//============================================================
// 文件: PLC_Logic.scl
// 项目: PLC-Robot-Integration-Demo (PLC控制ABB机器人码垛)
// 平台: TIA Portal V16+ / S7-1214C DC/DC/DC
// 内容: 伺服控制FB / 主顺控FB / 故障处理FB / 急停处理
// 版本: V2.3  日期: 2026-09-02
// 变更: V1.0 基础正反转+限位保护
//       V2.0 增加完整顺控、故障码、急停安全处理
//       V2.1 超时改锁存+定时器卫生(修超时后无法复位/误超时)
//            故障灯无故障时强制熄灭; 启动命令改600ms脉冲式;
//            满垛输出qRobotReset(DI2)通知机器人清垛位计数
//       V2.2 定时器实例声明由IEC_TIMER改为TON多重实例(IEC_TIMER是
//            定时器背景SDT, 不能按FB方式直接调用, "从源生成块"编译报错);
//            故障复位不再清nParts——机器人侧nCount(PERS)仅在满垛DI2时
//            清零, 两侧计数必须同步保持, 否则中垛复位后垛位错位且
//            PLC等满垛/机器人等DI2互等死锁
//       V2.3 bHomeDone/nParts/nPallet移入VAR RETAIN: 掉电重启后PLC侧
//            计数不再清零, 与机器人nCount(PERS)断电保持对齐, 堵住
//            断电重启失步入口(VAR RETAIN为IEC 61131-3标准声明段)
//============================================================
//
// ----------------- I/O 交叉引用表(调试用) -----------------
// I0.0 启动SB1(常开)      I0.1 停止SB2(常闭)
// I0.2 复位SB3            I0.3 手动/自动旋钮(自动=1)
// I0.4 正限位SQ1          I0.5 反限位SQ2
// I0.6 机器人"允许抓取"DO1 I0.7 物料检测光电E3Z
// I1.0 急停回路反馈(常闭)  I1.1 安全门开关(常闭)
// I1.2 机器人"码垛完成"DO2 I1.3 机器人故障DO3
// I1.4 伺服报警ALM(断=报警) I1.5 伺服就绪RDY
// Q0.0 脉冲PUL+  Q0.4 方向DIR+  Q0.3 伺服使能KA1
// Q0.1 运行绿灯 Q0.2 报警红灯  Q0.5 蜂鸣器    Q0.6 待机黄灯
// Q0.7 机器人DI1启动  Q1.0 机器人DI2复位
// MW10 电流  MW12 电压  MW14 温度  MW16 计数  MW22 故障码
// ----------------------------------------------------------
//============================================================

//============================================================
// 块1: FB_ServoCtrl —— 伺服使能/点动/限位保护/报警锁存
//============================================================
FUNCTION_BLOCK "FB_ServoCtrl"
{ S7_Optimized_Access := 'TRUE' }
VERSION: 1.0

VAR_INPUT
    bPowerOn    : BOOL;    // 使能命令(来自顺控或手动)
    bReset      : BOOL;    // 报警复位
    bJogFwd     : BOOL;    // 手动点动正转
    bJogRev     : BOOL;    // 手动点动反转
    bFwdLimit   : BOOL;    // 正向限位SQ1(1=压合)
    bRevLimit   : BOOL;    // 反向限位SQ2(1=压合)
    bServoReady : BOOL;    // 驱动器RDY(1=就绪)
    bServoFault : BOOL;    // 驱动器ALM(1=报警, 现场常闭取反后送入)
    bEStopOK    : BOOL;    // 急停回路(1=正常)
END_VAR

VAR_OUTPUT
    qEnable     : BOOL;    // 伺服使能 -> KA1 -> CN1.DI1(SON)
    qFwdAllow   : BOOL;    // 允许正转(软件许可)
    qRevAllow   : BOOL;    // 允许反转(软件许可)
    qRun        : BOOL;    // 运行中标志
    qAlarm      : BOOL;    // 伺服报警锁存输出
END_VAR

VAR
    bFaultLock  : BOOL;    // 故障锁存位
    iDiag       : INT;     // 诊断码(供HMI显示)
END_VAR

BEGIN
    //---- 1) 故障锁存: 报警或急停立即置位 ----
    IF bServoFault OR NOT bEStopOK THEN
        bFaultLock := TRUE;
        iDiag := 16#0101;              // 伺服报警/急停类
    END_IF;

    //---- 2) 双限位同时压合 = 接线故障, 同样锁存 ----
    IF bFwdLimit AND bRevLimit THEN
        bFaultLock := TRUE;
        iDiag := 16#0102;
    END_IF;

    //---- 3) 复位: 故障源消失后按复位才解锁 ----
    IF bReset AND NOT bServoFault AND bEStopOK
       AND NOT (bFwdLimit AND bRevLimit) THEN
        bFaultLock := FALSE;
        iDiag := 0;
    END_IF;

    //---- 4) 使能综合条件 ----
    qEnable := bPowerOn AND bServoReady
               AND NOT bFaultLock AND bEStopOK;

    //---- 5) 方向许可: 使能OK+未压限位+双命令互斥 ----
    qFwdAllow := qEnable AND NOT bFwdLimit
                 AND bJogFwd AND NOT bJogRev;
    qRevAllow := qEnable AND NOT bRevLimit
                 AND bJogRev AND NOT bJogFwd;

    qRun    := qFwdAllow OR qRevAllow;
    qAlarm  := bFaultLock;

END_FUNCTION_BLOCK


//============================================================
// 块2: FB_PalletMain —— 主顺控: 手动/自动/回原点/垛型计数
//============================================================
FUNCTION_BLOCK "FB_PalletMain"
{ S7_Optimized_Access := 'TRUE' }
VERSION: 2.0

VAR_INPUT
    bStart      : BOOL;    // 启动按钮I0.0
    bStop       : BOOL;    // 停止按钮I0.1(常闭,1=未按)
    bReset      : BOOL;    // 复位按钮I0.2
    bAutoSel    : BOOL;    // 自动模式I0.3(1=自动)
    bPartSeen   : BOOL;    // 物料检测I0.7
    bRobotAllow : BOOL;    // 机器人允许抓取DO1 -> I0.6
    bRobotDone  : BOOL;    // 码垛完成DO2 -> I1.2
    bRobotFault : BOOL;    // 机器人故障DO3 -> I1.3
    bEStopOK    : BOOL;    // 急停回路I1.0
    bDoorOK     : BOOL;    // 安全门I1.1
END_VAR

VAR_OUTPUT
    qServoPower : BOOL;    // 伺服使能命令(送FB_ServoCtrl)
    qRobotStart : BOOL;    // 机器人启动Q0.7->DI1
    qRobotReset : BOOL;    // 机器人复位Q1.0->DI2
    qLampRun    : BOOL;    // 运行绿灯
    qLampWait   : BOOL;    // 待机黄灯
    qLampFault  : BOOL;    // 故障红灯
    qBuzzer     : BOOL;    // 蜂鸣器
END_VAR

VAR
    iStep       : INT;     // 顺控步: 0待机 10回原点 20等料
                            // 30送料 40等允许 50发启动
                            // 60等完成 70垛满处理
    bStartPulse : BOOL;    // 启动按钮上升沿
    bStartMem   : BOOL;    // 启动边沿存储
    tonFeed     : TON;     // 送料超时监视(多重实例)
    tonHandShk  : TON;     // 握手超时监视(多重实例)
    tonBuzz     : TON;     // 蜂鸣限时(多重实例)
    tonStart    : TON;     // 启动命令脉宽控制(多重实例)
    bFeedTO     : BOOL;    // 送料超时锁存(复位前保持)
    bHandTO     : BOOL;    // 握手超时锁存(复位前保持)
    bAnyFault   : BOOL;    // 综合故障
END_VAR

VAR RETAIN
    bHomeDone   : BOOL;    // 原点完成标志(掉电保持)
    nParts      : INT;     // 本垛已码件数(掉电保持: 与机器人nCount(PERS)对齐,
                            // 否则断电后PLC清零而机器人保持, 垛位错位互等死锁)
    nPallet     : INT;     // 换垛计数(累计类, 掉电保持)
END_VAR

VAR CONSTANT
    cFeedTimeout  : TIME := T#8S;    // 送料超时(含物料堵塞)
    cHandTimeout  : TIME := T#30S;  // 机器人握手超时
    cBuzzTime     : TIME := T#3S;   // 报警蜂鸣时长
    cCmdPulse     : TIME := T#600MS; // 跨设备命令脉宽(防信号粘连)
    cPartsPerBox  : INT  := 48;     // 满垛件数 3x4x4
END_VAR

BEGIN
    //---- 1) 启动按钮上升沿 ----
    bStartPulse := bStart AND NOT bStartMem;
    bStartMem   := bStart;

    //---- 2) 综合故障 = 急停/门/机器人/超时锁存 ----
    // 超时用锁存位而非定时器Q直接参与: 定时器到点即复位,
    // 故障状态由锁存保持, 复位按钮清除, 避免"定时器残留导致
    // 无法复位"或"二次进入即超时"两类卡死
    bAnyFault := NOT bEStopOK OR NOT bDoorOK
                 OR bRobotFault OR bFeedTO OR bHandTO;

    //---- 3) 蜂鸣器: 故障瞬间响, 3秒后自停 ----
    tonBuzz(IN := bAnyFault, PT := cBuzzTime);
    qBuzzer := bAnyFault AND NOT tonBuzz.Q;

    //---- 4) 急停处理: 最高优先级, 立即撤使能与命令 ----
    IF bAnyFault THEN
        iStep        := 0;
        qServoPower  := FALSE;
        qRobotStart  := FALSE;
        qRobotReset  := FALSE;
        qLampRun     := FALSE;
        qLampWait    := FALSE;
        qLampFault   := TRUE;
        IF bReset AND bEStopOK AND bDoorOK AND NOT bRobotFault THEN
            // 复位: 故障源消失后清超时锁存。
            // 注意nParts不清零: 机器人nCount(PERS)仅在满垛经DI2清零,
            // 故障复位若单侧清零, 两侧对"第几件"失去共识——垛位换算
            // 错位, 且PLC永不满垛/机器人空等DI2, 互等30s超时死锁。
            // 两侧计数只能同步清零: 满垛换盘时PLC输出DI2, 机器人
            // 上升沿清nCount, PLC在步70按启动时清nParts。
            // 断电场景由VAR RETAIN保持nParts, 与nCount(PERS)对齐。
            bFeedTO := FALSE;
            bHandTO := FALSE;
        END_IF;
        RETURN;                          // 故障期间跳过顺控
    END_IF;

    qLampFault := FALSE;                 // 无故障时确保红灯熄灭

    //---- 5) 模式判断: 手动模式只允许伺服点动, 不发启动 ----
    IF NOT bAutoSel THEN
        iStep        := 0;
        qRobotStart  := FALSE;
        qRobotReset  := FALSE;
        qLampWait    := TRUE;
        qLampRun     := FALSE;
        qServoPower  := TRUE;            // 手动仍允许使能供点动
        RETURN;
    END_IF;

    //---- 6) 自动顺控状态机 ----
    IF NOT bStop THEN                    // 停止按钮(常闭断开)
        iStep := 0;
    END_IF;

    //---- 定时器卫生: 不属于对应步时强制复位 ----
    // 防止故障/停机打断后残留计时, 再次进入该步立即误超时
    IF iStep <> 30 THEN
        tonFeed(IN := FALSE);
    END_IF;
    IF NOT (iStep = 40 OR iStep = 60) THEN
        tonHandShk(IN := FALSE);
    END_IF;
    IF iStep <> 50 THEN
        tonStart(IN := FALSE);
    END_IF;

    CASE iStep OF

        0:  // 待机: 等待启动, 且必须先有原点
            qLampWait   := TRUE;
            qLampRun    := FALSE;
            qRobotStart := FALSE;
            IF bStartPulse THEN
                IF NOT bHomeDone THEN
                    iStep := 10;         // 先回原点
                ELSE
                    iStep := 20;
                END_IF;
            END_IF;

        10: // 回原点: 压SQ1后退回偏移量(此处由FB_Servo点动逻辑
            // 配合HMI手动完成, 自动回零用PTO回原点功能, 略)
            bHomeDone := TRUE;
            iStep     := 20;

        20: // 等料: 光电检测到物料进入送料步
            qServoPower := TRUE;
            qLampWait   := FALSE;
            qLampRun    := TRUE;
            IF bPartSeen THEN
                iStep := 30;
            END_IF;

        30: // 送料: 脉冲输出由Motion Control工艺对象完成,
            // 此处只做超时监视
            tonFeed(IN := TRUE, PT := cFeedTimeout);
            IF tonFeed.Q THEN
                bFeedTO := TRUE;         // 锁存送料超时, 进故障处理
                iStep   := 0;
            ELSIF NOT bPartSeen THEN     // 物料已离开检测位=送到位
                iStep := 40;
            END_IF;

        40: // 等机器人"允许抓取"
            tonHandShk(IN := TRUE, PT := cHandTimeout);
            IF bRobotAllow THEN
                iStep := 50;
            ELSIF tonHandShk.Q THEN
                bHandTO := TRUE;         // 锁存握手超时, 进故障处理
                iStep   := 0;
            END_IF;

        50: // 发启动命令(600ms脉冲式, 防信号粘连致机器人重复执行)
            qRobotStart := TRUE;
            tonStart(IN := TRUE, PT := cCmdPulse);
            IF tonStart.Q THEN           // 脉宽到, 撤命令进等待步
                iStep := 60;
            END_IF;

        60: // 等码垛完成(启动命令已在脉宽到点时撤除, 此处兜底清零)
            qRobotStart := FALSE;
            tonHandShk(IN := TRUE, PT := cHandTimeout);
            IF bRobotDone THEN
                nParts := nParts + 1;
                iStep  := 20;            // 下一件
            ELSIF tonHandShk.Q THEN
                bHandTO := TRUE;         // 锁存完成超时, 进故障处理
                iStep   := 0;
            END_IF;

        70: // 垛满: 提示换托盘(由完成计数触发进入)
            qLampWait    := TRUE;
            qLampRun     := FALSE;
            qServoPower  := FALSE;       // 换盘期间断开伺服使能
            // qRobotReset 保持输出, 机器人DI2上升沿清垛位计数
            IF bStartPulse THEN          // 换盘后按启动继续
                nParts       := 0;
                nPallet      := nPallet + 1;
                qRobotReset  := FALSE;   // 撤复位命令
                iStep        := 20;
            END_IF;

    END_CASE;

    IF nParts >= cPartsPerBox AND iStep = 20 THEN
        iStep       := 70;
        qRobotReset := TRUE;             // 满垛: 通知机器人准备新垛
    END_IF;

END_FUNCTION_BLOCK


//============================================================
// 块3: FB_FaultHandler —— 故障子程序: 优先级编码+首发故障锁存
// 注: 用FB而非FC, 静态变量才能跨周期保持"首发故障码"
//============================================================
FUNCTION_BLOCK "FB_FaultHandler"
{ S7_Optimized_Access := 'TRUE' }
VERSION: 1.0

VAR_INPUT
    bEStopOK    : BOOL;    // 1=正常
    bDoorOK     : BOOL;    // 1=正常
    bRobotFault : BOOL;    // 1=故障
    bServoFault : BOOL;    // 1=故障
    bFeedTO     : BOOL;    // 送料超时
    bHandTO     : BOOL;    // 握手超时
    bReset      : BOOL;    // 复位脉冲
END_VAR

VAR_OUTPUT
    wFaultCode  : WORD;    // 故障码(0=无故障, 供HMI显示)
    bFirstLock  : BOOL;    // 首发故障已锁存
END_VAR

VAR
    wCurrent    : WORD;    // 本周期按优先级算出的故障码
    wFirstCode  : WORD;    // 首发故障码(锁存)
END_VAR

BEGIN
    // 优先级: 急停 > 安全门 > 伺服 > 机器人 > 送料超时 > 握手超时
    IF NOT bEStopOK    THEN wCurrent := 16#0001;
    ELSIF NOT bDoorOK  THEN wCurrent := 16#0002;
    ELSIF bServoFault  THEN wCurrent := 16#0003;
    ELSIF bRobotFault  THEN wCurrent := 16#0004;
    ELSIF bFeedTO      THEN wCurrent := 16#0005;
    ELSIF bHandTO      THEN wCurrent := 16#0006;
    ELSE                    wCurrent := 16#0000;
    END_IF;

    // 首发故障锁存: 直到复位前保持不变, 便于现场定位
    IF wCurrent <> 16#0000 AND NOT bFirstLock THEN
        wFirstCode := wCurrent;
        bFirstLock := TRUE;
    END_IF;

    IF bReset AND wCurrent = 16#0000 THEN
        bFirstLock := FALSE;
        wFirstCode := 16#0000;
    END_IF;

    // 输出: 有故障显示当前码, 无故障时保留首发码(历史)供查询
    IF wCurrent <> 16#0000 THEN
        wFaultCode := wCurrent;
    ELSE
        wFaultCode := wFirstCode;
    END_IF;

END_FUNCTION_BLOCK

//============================================================
// OB1 调用示例(供参考, 在OB1中按如下方式接线):
//   CALL "FB_ServoCtrl", "FB_ServoCtrl_DB"
//        (bPowerOn:="FB_PalletMain_DB".qServoPower, ...)
//   CALL "FB_PalletMain", "FB_PalletMain_DB"
//        (bStart:="I0.0", bStop:="I0.1", ...)
//   CALL "FB_FaultHandler", "FB_FaultHandler_DB"
//        (bEStopOK:="I1.0",                       // 急停反馈
//         bFeedTO:="FB_PalletMain_DB".bFeedTO,
//         bHandTO:="FB_PalletMain_DB".bHandTO,
//         ... wFaultCode=>"MW22")
//============================================================
